FUNCTION_BLOCK "AnalogBatchProcessing"
VERSION : 0.1
BEGIN
END_FUNCTION_BLOCK
